(* CODESYS project 模拟量的分段线性标定(折线插值).library
   Author: Inovance
   Title: INOVANCE_Library
   Version: 0.0.0.0
   Placeholder: INOVANCE_Library
   DocFormat: reStructuredText
   DefaultNamespace: INOVANCE_Library
   Company: Inovance
   Description: Library For Demo

Project tree, tasks and I/O mapping:
  DataTypes/
    Enums/
    Structs/
    Alias/
    Unions/
  POUs/
    FunctionBlocks/
    Functions/
    Programs/
  GlobalVariables/
  Templates/
    data type STATE
    data type ERROR
    function block ETrig [ST]: prv_HandleDormantState, prv_HandleExecutingState, prv_HandleDoneState, prv_HandleErrorState, prv_HandleResettingState, pro_CyclicAction, pro_ResetAction
    function block LCon [ST]: prv_HandleDormantState, prv_HandleExecutingState, prv_HandleAbortingState, prv_HandleDoneState, prv_HandleErrorState, prv_HandleResettingState, pro_CyclicAction, pro_AbortAction, pro_ResetAction
    trigger_state_chart
    Level_state_detail
    Level_state_chart
    trigger_sequential
    trigger_state_detail
  00000000-0000-0000-0000-000000000000|C:\Users\r2317\Desktop\trigger_state_chart.png
  Interfaces/
  00000000-0000-0000-0000-000000000000|C:\Users\r2317\Desktop\Level_state_detail.png
  00000000-0000-0000-0000-000000000000|C:\Users\r2317\Desktop\Level_state_chart.png
  00000000-0000-0000-0000-000000000000|C:\Users\r2317\Desktop\trigger_sequential.png
  00000000-0000-0000-0000-000000000000|C:\Users\r2317\Desktop\trigger_state_detail.png
  program POU [ST]
*)

// Templates/STATE
{attribute 'qualified_only'}
{attribute 'strict'}
TYPE STATE :
(
	DORMANT, 	// Waiting for Start
	EXECUTING, 	// CyclicAction is running
	ABORTING,   // AbortAction is running
	DONE, 		// CyclicAction is complete
	ERROR, 		// Error condition reached
	RESETTING 	// ResetAction is running
);
END_TYPE

// Templates/ERROR
{attribute 'qualified_only'}
{attribute 'strict'}
TYPE ERROR :
(
	NO_ERROR :=0,
	TIME_OUT := 1
	(*...*)
);
END_TYPE

// Templates/ETrig
(* 
 * 这是最简单形式的功能，无论是文本还是图形表示，只有一个xExecute作为输入。为了描述这个FB的功能和行为，使用状态机图，描述不同的状态的结果转换。基本上有4种状态：休眠、忙碌、完成，结合重置和错误，见下图。
 *
 * .. image:: ../../Templates/trigger_state_chart.png
 *
 * 在输入xExecute检测到上升沿后，内部状态从休眠状态切换到忙状态，所有输入都被采样并存储，输出xBusy将设置为TRUE。 定义的操作将会启动，操作在运行过程中，会出现许多导致从Busy状态退出的条件，输出变量xBusy的值将设置为FALSE，内部状态机将从Busy切换到Done或Error状态之一。 
 * 此更改将镜像到输出变量xDone或xError之一。输出变量xBusy、xError、xDone互斥，同一时刻，只有一个输出变量为TRUE状态。
 * 
 * .. image:: ../../Templates/trigger_state_detail.png
 *
 * | Ready Condition: 如果操作已达到就绪状态而没有任何错误和时序错误，则输出变量xDone将设置为TRUE。内部状态从Busy切换到Done。
 * | Error Condition: 如果检测到错误条件，则输出变量xError设置为TRUE。内部状态从Busy切换到Error。此外，其中一个已定义的错误代码（本地枚举类型ERROR中的一个值）将分配给输出变量eError。
 *
 * 其中一个输出变量xDone或xError的值TRUE必须保持稳定最少一个周期。检测到输入变量xExecute的FALSE状态后，内部状态将切换为Reset。所有输出将初始化为其默认状态（重置输出）。  
 * 所有已声明的资源将被释放。 特别是输出变量xDone和xError将设置为FALSE。执行此重新初始化工作后，内部状态将从Reset切换到Dormant。
 *
 * 注意: 必须确保其中一个输出变量xDone或xError的状态TRUE必须保持稳定至少一个周期，例如添加子状态Sync。
 *
 * 下图是输入、输出状态和状态机时序图。
 *
 *  .. image:: ../../Templates/trigger_sequential.png
 *
 *)

FUNCTION_BLOCK ETrig
VAR_INPUT
	// Rising edge starts defined operation
	// FALSE => reset the defined operation
	// after ready condition was reached
	xExecute: BOOL;
END_VAR
VAR_OUTPUT
	// ready condition reached
	xDone: BOOL;
	// operation is running
	xBusy: BOOL;
	// error condition reached
	xError: BOOL;
	// error code describing error condition
	eErrorID : ERROR;
END_VAR

VAR
	eState : STATE;
	xFirstInvocation : BOOL := TRUE;
	xResetRequest : BOOL;
END_VAR

VAR_TEMP
	xAgain : BOOL;
END_VAR

REPEAT
	xAgain := FALSE;
	
	CASE eState OF
		STATE.DORMANT: 
			prv_HandleDormantState(xAgain=>xAgain);
			
		STATE.EXECUTING: 
			prv_HandleExecutingState(xAgain=>xAgain);
			
		STATE.DONE: 
			prv_HandleDoneState(xAgain=>xAgain);
			
		STATE.ERROR: 
			prv_HandleErrorState(xAgain=>xAgain);
			
		STATE.RESETTING: 
			prv_HandleResettingState(xAgain=>xAgain);
		
	END_CASE
	
UNTIL (NOT xAgain)
END_REPEAT;

METHOD PRIVATE prv_HandleDormantState
VAR_INPUT
END_VAR
VAR_OUTPUT 
	xAgain : BOOL; 
END_VAR
IF xExecute THEN 
	xBusy := TRUE; 
	eState := STATE.EXECUTING; 
	xAgain := TRUE; 
END_IF
END_METHOD

METHOD PRIVATE prv_HandleExecutingState
VAR_INPUT
END_VAR
VAR_OUTPUT 
	xAgain : BOOL; 
END_VAR 
VAR 
	xComplete : BOOL; 
END_VAR
pro_CyclicAction( xComplete=>xComplete, eErrorID=>eErrorID );
IF eErrorID <> ERROR.NO_ERROR THEN 
	eState := STATE.ERROR; 
	xAgain := TRUE;
ELSIF xComplete THEN 
	eState := STATE.DONE; 
	xAgain := TRUE; 
END_IF
END_METHOD

METHOD PRIVATE prv_HandleDoneState
VAR_INPUT
END_VAR
VAR_OUTPUT 
	xAgain : BOOL; 
END_VAR
IF xDone AND (xResetRequest OR NOT xExecute) THEN 
	eState := STATE.RESETTING; 
	xAgain := TRUE;
ELSE 
	xBusy := FALSE; 
	xDone := TRUE; 
	xResetRequest := NOT xExecute; 
	xAgain := FALSE; (* !!! *) 
END_IF
END_METHOD

METHOD PRIVATE prv_HandleErrorState
VAR_INPUT
END_VAR
VAR_OUTPUT 
	xAgain : BOOL; 
END_VAR
IF xError AND (xResetRequest OR NOT xExecute) THEN 
	eState := STATE.RESETTING; 
	xAgain := TRUE;
ELSE 
	xBusy := FALSE; 
	xError := TRUE; 
	xResetRequest := NOT xExecute;
	xAgain := FALSE; (* !!! *) 
END_IF
END_METHOD

METHOD PRIVATE prv_HandleResettingState
VAR_INPUT
END_VAR
VAR_OUTPUT 
	xAgain : BOOL; 
END_VAR 
VAR 
	xComplete : BOOL; 
END_VAR
pro_ResetAction(xComplete=>xComplete); 
IF xComplete THEN 
	xBusy := FALSE; 
	xDone := FALSE; 
	xError := FALSE; 
	eErrorID := ERROR.NO_ERROR; 
	eState := STATE.DORMANT; 
	xFirstInvocation := TRUE; 
	xAgain := xResetRequest; (* !!! *) 
	xResetRequest := FALSE; 
END_IF
END_METHOD

METHOD PROTECTED pro_CyclicAction
VAR_INPUT
END_VAR
VAR_OUTPUT 
	xComplete : BOOL;
	eErrorID : ERROR; 
END_VAR
IF xFirstInvocation THEN 
	(* Starting *) 
    // for the first (!) invocation, 
	// sample the input variables 
	xFirstInvocation := FALSE; 
END_IF

(* Executing *)
// working to reach the ready condition 
// => xComplete := TRUE 
// if an error condition is reached 
// => set eErrorID to a value other than ERROR.NO_ERROR 

xComplete := TRUE; 
eErrorID := ERROR.NO_ERROR; 

IF xComplete OR eErrorID <> ERROR.NO_ERROR THEN 
	(* Cleaning *) 
	// if possible free as much allocated resources
	// as possible 
END_IF
END_METHOD

METHOD PROTECTED pro_ResetAction
VAR_INPUT
END_VAR
VAR_OUTPUT 
	xComplete : BOOL; 
END_VAR
// free all allocated resources 
// reinitialize instance variables 
xComplete := TRUE;
END_METHOD

END_FUNCTION_BLOCK

// Templates/LCon
(*
 * 此状态图包含5种状态：休眠，执行，完成，错误和中止，但为了清楚起见，在图中添加了一个重置状态.
 *
 * .. image:: ../../Templates/Level_state_chart.png
 *
 * 在输入xEnable检测到上升沿后，内部状态从休眠状态切换到忙状态，所有输入都被采样并存储，输出xBusy将设置为TRUE。定义的操作将会启动，操作在运行过程中，会出现许多导致从Busy状态退出的条件，输出变量xBusy的值将设置为FALSE，内部状态机将从Busy切换到Done或Error状态之一。
 * 
 * 此更改将镜像到输出变量xDone或xError之一。输出变量xBusy、xError、xDone互斥，同一时刻，只有一个输出变量为TRUE状态。
 * 
 *  .. image:: ../../Templates/Level_state_detail.png
 * 
 * 有些使用场合，xDone被xValid替换，或者没有xDone，具体内容参考标准《PLCopen Software Creation Guidelines:Creating PLCopen Compliant Libraries》，该标准详细描述了边沿控制、电平控制分类，输入、输出、状态机、实现代码，功能块集合， 
 *)


FUNCTION_BLOCK LCon
VAR_INPUT
	// TRUE => activate the defined operation
	// FALSE => abort/reset the defined operation
	xEnable: BOOL;
END_VAR
VAR_OUTPUT
	// ready condition reached
	xDone: BOOL;  
	// operation is running
	xBusy: BOOL;
	// error condition reached
	xError: BOOL;
	// error code describing error conditions
	eErrorID : ERROR;
END_VAR

VAR
	eState : STATE;
	xResetRequest : BOOL;
END_VAR

VAR_TEMP
	xAgain : BOOL;
END_VAR

REPEAT
	xAgain := FALSE;
	
	CASE eState OF
		STATE.DORMANT: 
			prv_HandleDormantState(xAgain=>xAgain);
			
		STATE.EXECUTING: 
			prv_HandleExecutingState(xAgain=>xAgain);
			
		STATE.DONE: 
			prv_HandleDoneState(xAgain=>xAgain);
			
		STATE.ERROR: 
			prv_HandleErrorState(xAgain=>xAgain);
			
		STATE.ABORTING: 
			prv_HandleAbortingState(xAgain=>xAgain);
			
		STATE.RESETTING: 
			prv_HandleResettingState(xAgain=>xAgain);
	END_CASE
	
UNTIL (NOT xAgain)
END_REPEAT;

METHOD PRIVATE prv_HandleDormantState
VAR_INPUT
END_VAR
VAR_OUTPUT 
	xAgain : BOOL; 
END_VAR
IF xEnable THEN 
	xBusy := TRUE; 
	eState := STATE.EXECUTING; 
	xAgain := TRUE; 
END_IF
END_METHOD

METHOD PRIVATE prv_HandleExecutingState
VAR_INPUT
END_VAR
VAR_OUTPUT 
	xAgain : BOOL; 
END_VAR 
VAR 
	xComplete : BOOL; 
	xTimeOut : BOOL;
END_VAR
IF xEnable THEN
	pro_CyclicAction( xComplete=>xComplete, eErrorID=>eErrorID );
END_IF

IF eErrorID <> ERROR.NO_ERROR THEN 
	eState := STATE.ERROR; 
	xAgain := TRUE;
ELSIF NOT xEnable THEN
	eState := STATE.ABORTING;
	xAgain := TRUE;
ELSIF xComplete THEN 
	eState := STATE.DONE; 
	xAgain := TRUE; 
END_IF
END_METHOD

METHOD PRIVATE prv_HandleAbortingState
VAR_INPUT
END_VAR
VAR_OUTPUT 
	xAgain : BOOL; 
END_VAR 
VAR 
	xComplete : BOOL; 
END_VAR
pro_AbortAction( xComplete=>xComplete, eErrorID=>eErrorID );
IF eErrorID <> ERROR.NO_ERROR THEN
	eState := STATE.ERROR; 
	xAgain := TRUE;
	
ELSIF xComplete THEN
	eState := STATE.RESETTING;
	xAgain := TRUE;
END_IF
END_METHOD

METHOD PRIVATE prv_HandleDoneState
VAR_INPUT
END_VAR
VAR_OUTPUT 
	xAgain : BOOL; 
END_VAR
IF xDone AND NOT xEnable THEN 
	eState := STATE.RESETTING; 
	xAgain := TRUE;
ELSE 
	xBusy := FALSE; 
	xDone := TRUE; 
	xAgain := FALSE; (* !!! *) 
END_IF
END_METHOD

METHOD PRIVATE prv_HandleErrorState
VAR_INPUT
END_VAR
VAR_OUTPUT 
	xAgain : BOOL; 
END_VAR
IF xError AND (xResetRequest OR NOT xEnable) THEN 
	eState := STATE.RESETTING;
	xAgain := TRUE;
ELSE 
	xBusy := FALSE; 
	xError := TRUE; 
	xResetRequest := NOT xEnable;
	xAgain := FALSE; (* !!! *) 
END_IF
END_METHOD

METHOD PRIVATE prv_HandleResettingState
VAR_INPUT
END_VAR
VAR_OUTPUT 
	xAgain : BOOL; 
END_VAR 
VAR 
	xComplete : BOOL; 
END_VAR
pro_ResetAction(xComplete=>xComplete); 
IF xComplete THEN 
	xBusy := FALSE; 
	xDone := FALSE; 
	xError := FALSE; 
	eErrorID := ERROR.NO_ERROR; 
	eState := STATE.DORMANT; 
	xAgain := xResetRequest; (* !!! *) 
	xResetRequest := FALSE; 
END_IF
END_METHOD

METHOD PROTECTED pro_CyclicAction
VAR_INPUT
END_VAR
VAR_OUTPUT 
	xComplete : BOOL;
	eErrorID : ERROR; 
END_VAR
IF xEnable THEN 
	(* Executing *)
	// for every invocation, 
	// sample the input variables 
	// working to reach the ready condition 
	// ⇒ xComplete := TRUE 
	// if an error condition is reached set 
	// eErrorID to a value other than ERROR.NO_ERROR
	
	xComplete := TRUE; 
	eErrorID := ERROR.NO_ERROR; 	
END_IF


IF NOT xEnable OR xComplete OR eErrorID <> ERROR.NO_ERROR THEN
	(* Cleaning *) 
	// if possible free as much allocated resources
	// as possible 
END_IF
END_METHOD

METHOD PROTECTED pro_AbortAction
VAR_INPUT
END_VAR
VAR_OUTPUT 
	xComplete : BOOL;
	eErrorID : ERROR; 
END_VAR
// abort all running operations 
// if an error condition is reached set 
// eErrorID to a value other than ERROR.NO_ERROR 

xComplete := TRUE;
eErrorID := ERROR.NO_ERROR;
END_METHOD

METHOD PROTECTED pro_ResetAction
VAR_INPUT
END_VAR
VAR_OUTPUT 
	xComplete : BOOL; 
END_VAR
// free all allocated resources 
// reinitialize instance variables 
xComplete := TRUE;
END_METHOD

END_FUNCTION_BLOCK

// POU
PROGRAM POU
VAR_INPUT
	real_D_now:INT;
	real_D:ARRAY[1..10] OF INT;
	test_D:ARRAY[1..10]  OF INT;
END_VAR
VAR_OUTPUT
	out_D:INT;
END_VAR
VAR
	n:INT;
	ratio:ARRAY[1..10] OF REAL;
	point_1:INT;
END_VAR

//功能1，对曲线进行修正后，将当前值换算后输出。
//功能2，如果输入值突变，进行累加变化，达到目标值,如何实现？监测突变、突变则执行程序，进行输出规划，并按照既定规划进行输出。
//point判断，防止计算错误
point_1:=10;
//计算每段折线的斜率
FOR n:=1 TO point_1-1 DO
	ratio[n]:=INT_TO_REAL(real_D[n+1]-real_D[n])/INT_TO_REAL(test_D[n+1]-test_D[n]);
END_FOR
//计算输入值在区间内时的输出结果
FOR n:=1 TO point_1-1 DO
    IF real_D_now>real_D[n] AND real_D_now<real_D[n+1] THEN
		real_D_now:=real_D[n]+REAL_TO_INT((real_D_now-real_D[n])/ratio[n]);
    END_IF
END_FOR
//计算输入值小于区间内时的输出结果
IF real_D_now<real_D[1] THEN
	real_D_now:=test_D[1]-REAL_TO_INT(INT_TO_REAL(real_D[n]-real_D_now)/ratio[1]);
END_IF
//计算输入值大于区间内时的输出结果
IF real_D_now >= real_D [point_1] THEN
	out_D := test_D[point_1] +REAL_TO_INT ( INT_TO_REAL  (real_D_now - real_D[ point_1] )/ ratio[point_1-1]);
END_IF;

END_PROGRAM
